(* PLC project opcua_server, Beremiz opcua_server 1 *)
(* stored: creationDateTime 2026-10-11T12:00:00, modificationDateTime 2026-10-11T12:00:00 *)

TYPE POINT : STRUCT
  X : INT;
  Y : REAL;
END_STRUCT;
END_TYPE

FUNCTION_BLOCK COUNTER_FB
  VAR_OUTPUT
    CNT : DINT;
  END_VAR

            CNT := CNT + 1;
          
END_FUNCTION_BLOCK

PROGRAM program0
  VAR
    Counter : COUNTER_FB;
    Arr : ARRAY[0..2] OF INT;
    Pt : POINT;
    Pts : ARRAY[1..2] OF POINT;
    Cmd : INT;
    Echo : INT;
    Msg : STRING := 'hello';
    Delay : TIME := T#1500ms;
    LOGGER0 : LOGGER;
  END_VAR
  VAR_EXTERNAL
    GFlag : BOOL;
  END_VAR

            Counter();
Arr[1] := Arr[0] * 2;
Pts[2].X := Pt.X + 1;
IF Cmd <> Echo THEN
  Echo := Cmd;
  LOGGER0(TRIG := TRUE, MSG := CONCAT('OPCUA write Cmd=', INT_TO_STRING(Cmd)));
ELSE
  LOGGER0(TRIG := FALSE);
END_IF;
          
END_PROGRAM

CONFIGURATION config
  VAR_GLOBAL
    GFlag : BOOL;
  END_VAR
  RESOURCE resource1 ON PLC
    VAR_GLOBAL
      RVar : DINT;
    END_VAR
    TASK task0(INTERVAL := T#100ms, PRIORITY := 0);
    PROGRAM instance0 WITH task0 : program0;
  END_RESOURCE
END_CONFIGURATION
